FUNCTION_BLOCK fbShutterCmdSourceSwitch IMPLEMENTS iShutterCmdSource
VAR_INPUT
    OpenSwitchState : stSwitchState;
    CloseSwitchState : stSwitchState;
    ShutterStateType : eShutterStateType;
	ShutterConfig : stShutterConfig;
END_VAR

METHOD Process
VAR_IN_OUT
	CmdEvent : stShutterCmdEvent;
END_VAR

// Exit if both switches are idle
IF OpenSwitchState.StateType = eSwitchStateType.IDLE AND
   CloseSwitchState.StateType = eSwitchStateType.IDLE THEN
    RETURN;
END_IF

// If shutter is moving and any switch was pressed
IF ShutterStateType <> eShutterStateType.IDLE THEN
    CmdEvent.Cmd.CmdType := eShutterCmdType.STOP;
// Double Open click
ELSIF (OpenSwitchState.StateType = eSwitchStateType.MULTI_CLICK) AND (OpenSwitchState.PressCount = 2) THEN
    CmdEvent.Cmd.CmdType := eShutterCmdType.OPEN;
// Double Close click
ELSIF (CloseSwitchState.StateType = eSwitchStateType.MULTI_CLICK) AND (CloseSwitchState.PressCount = 2) THEN
    CmdEvent.Cmd.CmdType := eShutterCmdType.CLOSE;
// Triple Open click
ELSIF (OpenSwitchState.StateType = eSwitchStateType.MULTI_CLICK) AND (OpenSwitchState.PressCount = 3) THEN
    CmdEvent.Cmd.CmdType := eShutterCmdType.SAVE_POS1;
// Triple Close click
ELSIF (CloseSwitchState.StateType = eSwitchStateType.MULTI_CLICK) AND (CloseSwitchState.PressCount = 3) THEN
    CmdEvent.Cmd.CmdType := eShutterCmdType.SAVE_POS2;
// Short Open click
ELSIF OpenSwitchState.StateType = eSwitchStateType.SHORT_CLICK THEN
    CmdEvent.Cmd.CmdType := eShutterCmdType.STEP_OPEN;
// Short Close click
ELSIF CloseSwitchState.StateType = eSwitchStateType.SHORT_CLICK THEN
    CmdEvent.Cmd.CmdType := eShutterCmdType.STEP_CLOSE;
// Long Open click
ELSIF OpenSwitchState.StateType = eSwitchStateType.LONG_CLICK THEN
    CmdEvent.Cmd.CmdType := eShutterCmdType.MOVE_TO_POSITION;
    CmdEvent.Cmd.Position := ShutterConfig.SavedPosition1;
// Long Close click
ELSIF CloseSwitchState.StateType = eSwitchStateType.LONG_CLICK THEN
    CmdEvent.Cmd.CmdType := eShutterCmdType.MOVE_TO_POSITION;
    CmdEvent.Cmd.Position := ShutterConfig.SavedPosition2;
END_IF

CmdEvent.Execute := TRUE;
CmdEvent.Source := eShutterCmdSource.SWITCH;
END_METHOD

END_FUNCTION_BLOCK

(* stored: Version 1.1.0.1
   POU fbShutterCmdSourceSwitch: Id {c862dcf9-c651-483d-a78a-0c62d3a73fd7}, SpecialFunc None
   Method Process: Id {bb7c2f45-924d-4762-a2d7-89765f3d0a73} *)
